TYPE E_State :
(
  Idle,
  Busy
);
END_TYPE

(* stored: Version 1.1.0.1
   DUT E_State: Id {00000000-0000-0000-0000-000000000002} *)
